// Réponse de l'opérateur (docs/06 § 6.2) ; nStation 0 = calibration machine
{attribute 'pack_mode' := '1'}
TYPE ST_PromptAnswer :
STRUCT
    nSeq : UDINT;
    nStation : USINT;
    nPromptId : UDINT;
    bConfirm : BOOL;                // faux = annuler
    fValue : LREAL;
    sUser : STRING(24);
END_STRUCT
END_TYPE

(* stored: Version 1.1.0.1, ProductVersion 3.1.4024.12
   DUT ST_PromptAnswer: Id {8b2aff6b-e179-5d9f-bff8-940cb0499cfe} *)
